Fanuc KAREL source: kt00901.KL

-- PROVISIONAL review KL for V1013-1; original PC SHA256 38f2757c90a8aa9ad6170158dc6b63b7d40590818b72a7560a5d1180666ff95b
-- Incomplete behavior may be omitted. Consult companion uncertainty JSON. Do not deploy.
PROGRAM KT00901
%NOLOCKGROUP
VAR
  OUT : BOOLEAN
-- UNRESOLVED_DECL P1 type=000199
-- UNRESOLVED_DECL P2 type=000199
BEGIN
  -- UNRESOLVED_PC offsets 5-28; opcodes 27,22,1C,27,9D,76,23
  -- UNRESOLVED_PC offsets 33-37; opcodes 7F
END KT00901
